Fanuc KAREL source: kd00052.KL

-- PROVISIONAL review KL for V1013-1; original PC SHA256 37b30c328d807954e4dd12ede16a00a1f23a8f5bb997ccf6639d6386f61c69be
-- Incomplete behavior may be omitted. Consult companion uncertainty JSON. Do not deploy.
PROGRAM KD00052
%NOLOCKGROUP
VAR
  I : INTEGER
  J : INTEGER
  B : BOOLEAN
  R : REAL
  S : STRING[80]
-- UNRESOLVED_DECL P type=000101
BEGIN
  -- UNRESOLVED_PC offsets 5-42; opcodes 01,22,1C,06,82,03,9D,2E,51,9D,12,9D,1B,9D,13,04,0B
  -- UNRESOLVED_PC offsets 47-51; opcodes 7F
END KD00052
